(* Logix 5000 project; controller TFF vendor 1 type 14 code 107 rev 34.11; software revision 34.03; part 25 of 36 *)
(* tags used below, declared in another part *)
   Address : DINT;   // Temp Address
   Index : DINT;   // Index
   PCV101_PID_Settings : INT;
   sBar1 : STRING5;
   sBar2 : STRING5;
   sBar3 : STRING5;
   AnalogOutput : AnalogOutput[25];   // Analog Output Array
   Concentration : Concentration;
   ControlLoop_FeedBagLevel : ALIAS FOR ControlLoop[2];   // Feed Bag Level Control Loop
   ControlLoop_FeedPump : ALIAS FOR ControlLoop[1];   // Feed Pump Control Loop
   ControlLoop_PCV101 : ALIAS FOR ControlLoop[5];   // PCV101 Control Loop
   ControlLoop_PCV101_5ms : ALIAS FOR ControlLoop[6];   // PCV101 Control Loop
   ControlLoop_PCV101_CV : REAL;   // Control Value
   ControlLoop_PCV101_RAMP_OUT : REAL;   // Ramp Output
   DerivedData : DerivedData;   // Derived data (user input and calculated values)
   Diafiltration : Diafiltration;
   DigitalOutput : BOOL[256];   // Digital Output Array these bits are sent to output cards.
   DigitalPoint : DigitalPoint[150];   // Digital Point Array
   DP : ALIAS FOR AnalogPoint[40];   // Differential Pressure
   DPAlarm : ALIAS FOR AlarmAnalog[40];   // Differential Pressure Alarm
   Drive : Drive[11];   // Drives Array
   FI001 : ALIAS FOR AnalogPoint[42];   // Feed Flow
   FI001Alarm : ALIAS FOR AlarmAnalog[42];   // Feed Flow Alarm
   FI003 : ALIAS FOR AnalogPoint[17];
   FI101 : ALIAS FOR AnalogPoint[2];   // Filtrate Flow
   FI401 : ALIAS FOR AnalogPoint[43];   // Transfer Pump Flow
   FI401Alarm : ALIAS FOR AlarmAnalog[43];   // Transfer Pump Flow Alarm
   FlowPath : FlowPath[64];   // Flow Path Array
   FlowPathControl : FlowPathControl;   // Flow Path Control
   FQ_Conc : ALIAS FOR Totalizer[0];   // Concentration Totalizer
   FQ_Diaf : ALIAS FOR Totalizer[1];   // DiafiltrationTotalizer
   LI001 : ALIAS FOR AnalogPoint[44];   // Feed Bag Volume
   Membrane_Data : Membrane_Data;   // Membrane Data
   NWP : ALIAS FOR AnalogPoint[45];   // Normalized Water Permeability
   Options : Options;   // Options List
   PCV101_Control : PCV_Control;   // PCV101 Control UDT
   PERM : ALIAS FOR AnalogPoint[46];   // Membrane Permeability
   Phase : Phases[6];   // Phase Control Array
   Phase0 : ALIAS FOR Phase[0];   // Phase 0
   PhaseTotalizer : PhaseTotalizer[18];   // Phase Totalizers Array
   PI001 : ALIAS FOR AnalogPoint[5];   // Feed Pressure
   PI002 : ALIAS FOR AnalogPoint[6];   // Retentate Pressure
   PI101 : ALIAS FOR AnalogPoint[7];   // Filtrate Pressure
   PI401 : ALIAS FOR AnalogPoint[8];   // Transfer Pump Pressure
   PipeAnimation : PipeAnimation;   // HMI Pipe Animation Array
   SIC001 : ALIAS FOR Drive[1];   // Feed Pump
   SIC001DF : ALIAS FOR DigitalPoint[8];   // Feed Pump Defect
   SIC002 : ALIAS FOR Drive[2];   // Transfer Pump
   SIC002DF : ALIAS FOR DigitalPoint[9];   // Transfer Pump Defect
   SysControl : SysControl;   // General system status and command
   ThisSystem : SystemType;
   TI001 : ALIAS FOR AnalogPoint[13];   // Feed Bag Temperature
   TMP : ALIAS FOR AnalogPoint[41];   // Trans-membrane Pressure
   TMPAlarm : ALIAS FOR AlarmAnalog[41];   // Trans-membrane Pressure Alarm
   Totalizer : Totalizers[20];   // Totalizers Array
   XS011 : ALIAS FOR DigitalPoint[11];   // Pump P001 Type
   XS012 : ALIAS FOR DigitalPoint[12];   // Pump P002 Type
(* Process, continued *)

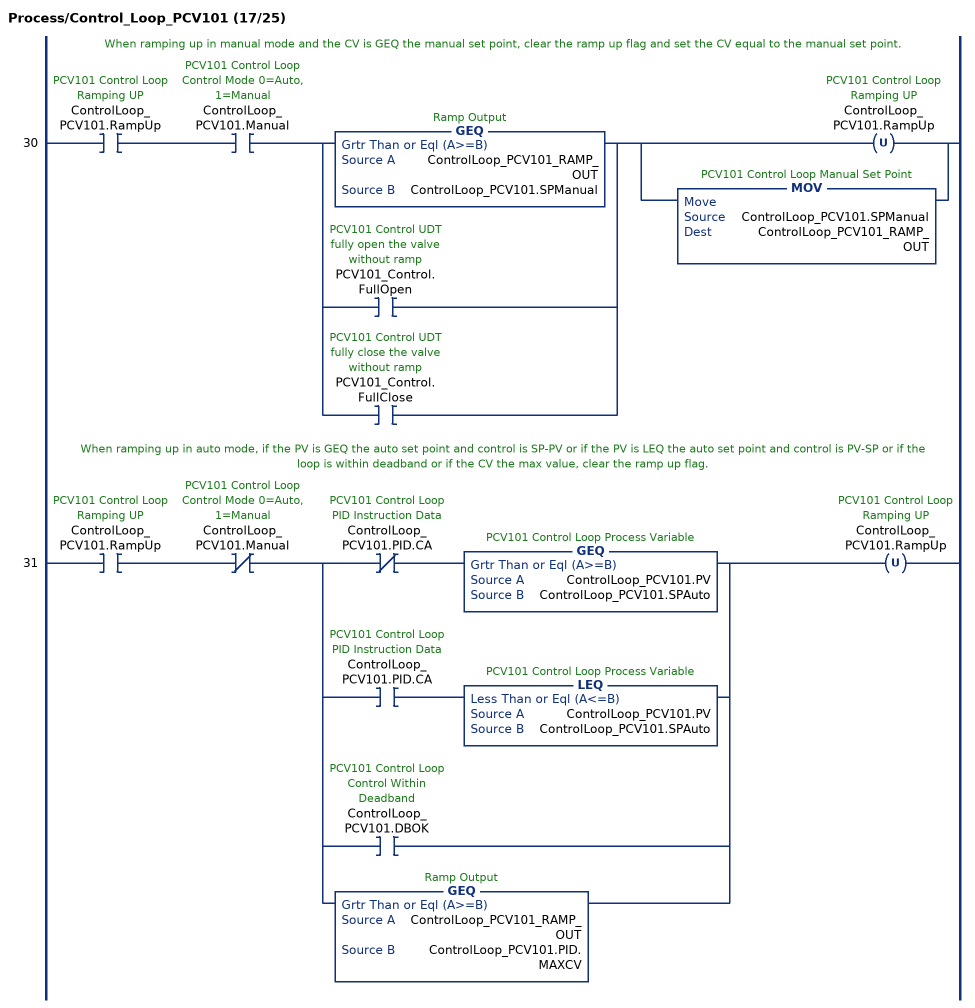
   [picture p237: Process/Control_Loop_PCV101 rungs 30-31]
   // When ramping up in manual mode and the CV is GEQ the manual set point, clear the ramp up flag and set the CV equal to the manual set point.
   30: XIC(ControlLoop_PCV101.RampUp)XIC(ControlLoop_PCV101.Manual)[GEQ(ControlLoop_PCV101_RAMP_OUT,ControlLoop_PCV101.SPManual) ,XIC(PCV101_Control.FullOpen) ,XIC(PCV101_Control.FullClose) ][OTU(ControlLoop_PCV101.RampUp) ,MOV(ControlLoop_PCV101.SPManual,ControlLoop_PCV101_RAMP_OUT) ];
   // When ramping up in auto mode, if the PV is GEQ the auto set point and control is SP-PV or if the PV is LEQ the auto set point and control is PV-SP or if the loop is within deadband or if the CV the max value, clear the ramp up flag.
   31: XIC(ControlLoop_PCV101.RampUp)XIO(ControlLoop_PCV101.Manual)[XIO(ControlLoop_PCV101.PID.CA) GEQ(ControlLoop_PCV101.PV,ControlLoop_PCV101.SPAuto) ,XIC(ControlLoop_PCV101.PID.CA) LEQ(ControlLoop_PCV101.PV,ControlLoop_PCV101.SPAuto) ,XIC(ControlLoop_PCV101.DBOK) ,GEQ(ControlLoop_PCV101_RAMP_OUT,ControlLoop_PCV101.PID.MAXCV) ]OTU(ControlLoop_PCV101.RampUp);
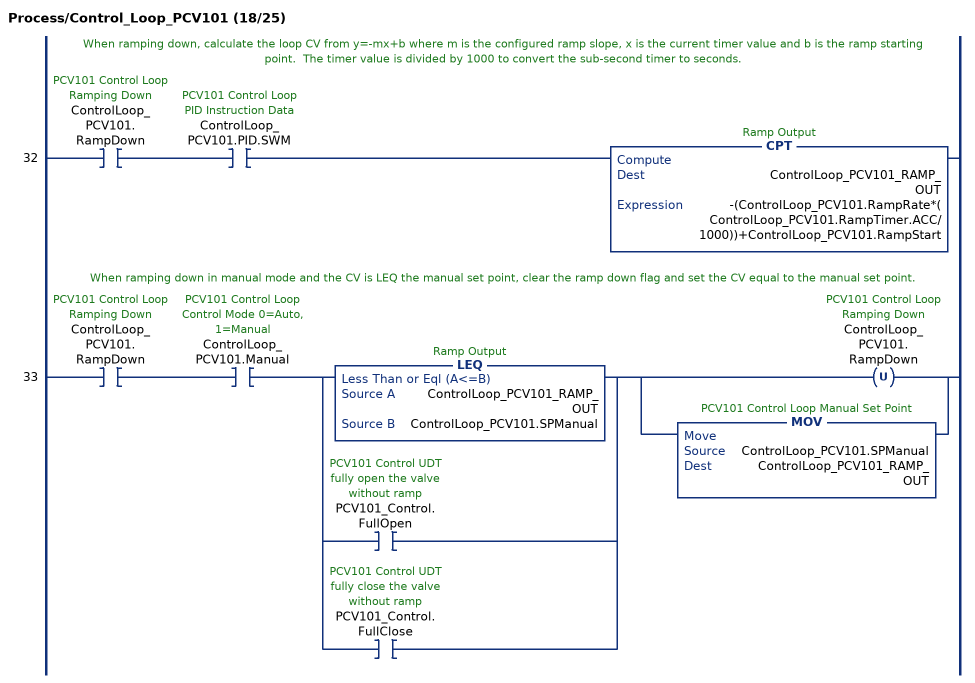
   // When ramping down, calculate the loop CV from y=-mx+b where m is the configured ramp slope, x is the current timer value and b is the ramp starting point.  The timer value is divided by 1000 to convert the sub-second timer to seconds.
   32: XIC(ControlLoop_PCV101.RampDown)XIC(ControlLoop_PCV101.PID.SWM)CPT(ControlLoop_PCV101_RAMP_OUT,-(ControlLoop_PCV101.RampRate*(ControlLoop_PCV101.RampTimer.ACC/1000))+ControlLoop_PCV101.RampStart);
   // When ramping down in manual mode and the CV is LEQ the manual set point, clear the ramp down flag and set the CV equal to the manual set point.
   33: XIC(ControlLoop_PCV101.RampDown)XIC(ControlLoop_PCV101.Manual)[LEQ(ControlLoop_PCV101_RAMP_OUT,ControlLoop_PCV101.SPManual) ,XIC(PCV101_Control.FullOpen) ,XIC(PCV101_Control.FullClose) ][OTU(ControlLoop_PCV101.RampDown) ,MOV(ControlLoop_PCV101.SPManual,ControlLoop_PCV101_RAMP_OUT) ];
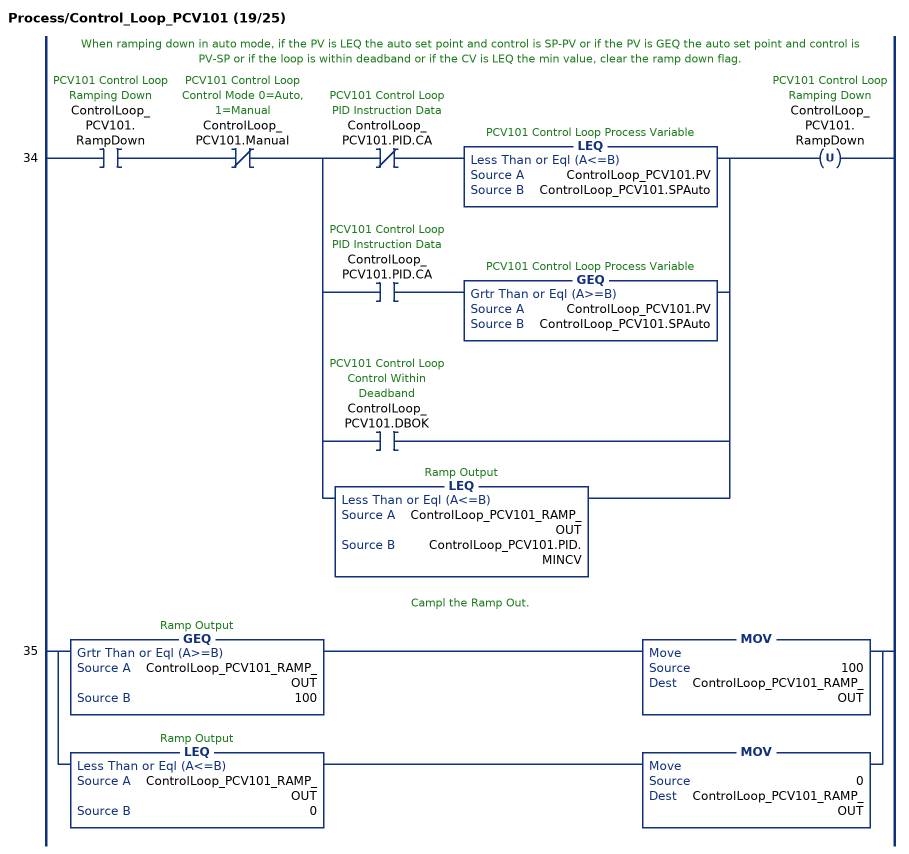
   // When ramping down in auto mode, if the PV is LEQ the auto set point and control is SP-PV or if the PV is GEQ the auto set point and control is PV-SP or if the loop is within deadband or if the CV is LEQ the min value, clear the ramp down flag.
   34: XIC(ControlLoop_PCV101.RampDown)XIO(ControlLoop_PCV101.Manual)[XIO(ControlLoop_PCV101.PID.CA) LEQ(ControlLoop_PCV101.PV,ControlLoop_PCV101.SPAuto) ,XIC(ControlLoop_PCV101.PID.CA) GEQ(ControlLoop_PCV101.PV,ControlLoop_PCV101.SPAuto) ,XIC(ControlLoop_PCV101.DBOK) ,LEQ(ControlLoop_PCV101_RAMP_OUT,ControlLoop_PCV101.PID.MINCV) ]OTU(ControlLoop_PCV101.RampDown);
   // Campl the Ramp Out.
   35: [GEQ(ControlLoop_PCV101_RAMP_OUT,100) MOV(100,ControlLoop_PCV101_RAMP_OUT) ,LEQ(ControlLoop_PCV101_RAMP_OUT,0) MOV(0,ControlLoop_PCV101_RAMP_OUT) ];
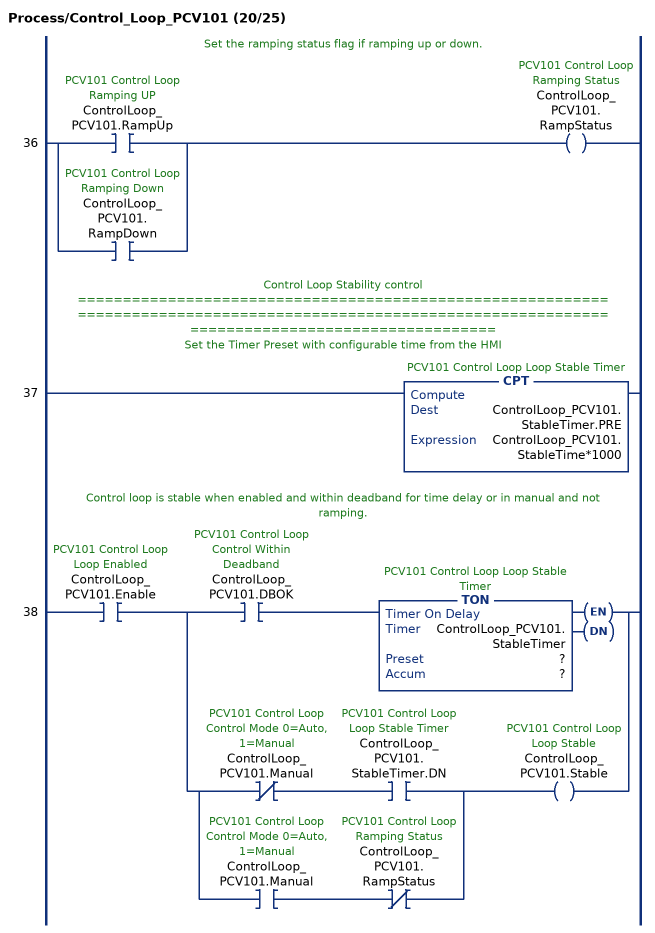
   // Set the ramping status flag if ramping up or down.
   36: [XIC(ControlLoop_PCV101.RampUp) ,XIC(ControlLoop_PCV101.RampDown) ]OTE(ControlLoop_PCV101.RampStatus);
   // Control Loop Stability control
   // ========================================================================================================================================================
   // Set the Timer Preset with configurable time from the HMI
   37: CPT(ControlLoop_PCV101.StableTimer.PRE,ControlLoop_PCV101.StableTime*1000);
   // Control loop is stable when enabled and within deadband for time delay or in manual and not ramping.
   38: XIC(ControlLoop_PCV101.Enable)[XIC(ControlLoop_PCV101.DBOK) TON(ControlLoop_PCV101.StableTimer,?,?) ,[XIO(ControlLoop_PCV101.Manual) XIC(ControlLoop_PCV101.StableTimer.DN) ,XIC(ControlLoop_PCV101.Manual) XIO(ControlLoop_PCV101.RampStatus) ] OTE(ControlLoop_PCV101.Stable) ];
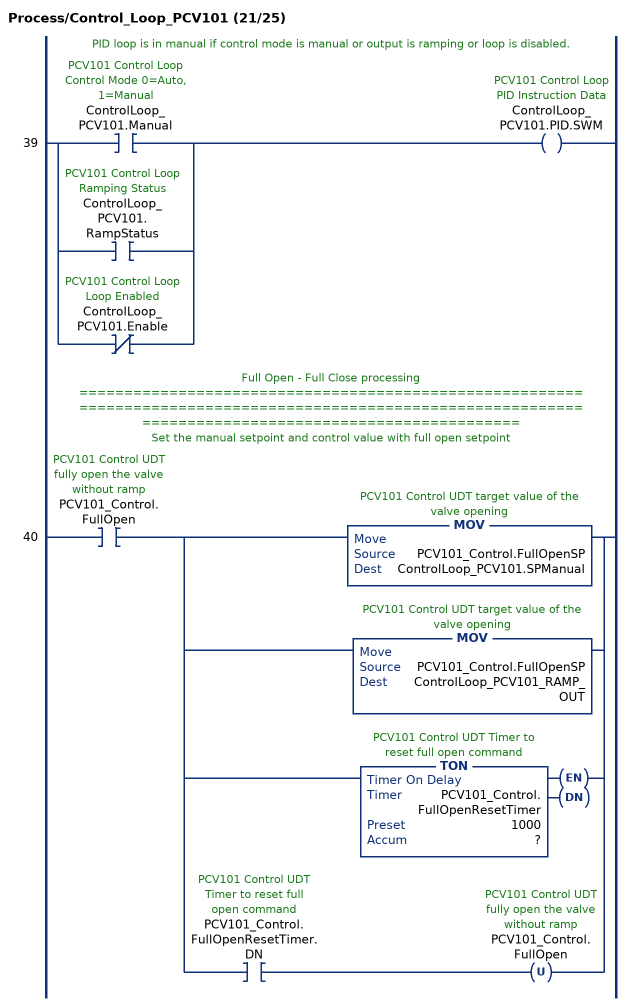
   // PID loop is in manual if control mode is manual or output is ramping or loop is disabled.
   39: [XIC(ControlLoop_PCV101.Manual) ,XIC(ControlLoop_PCV101.RampStatus) ,XIO(ControlLoop_PCV101.Enable) ]OTE(ControlLoop_PCV101.PID.SWM);
   // Full Open - Full Close processing
   // ==========================================================================================================================================================
   // Set the manual setpoint and control value with full open setpoint
   40: XIC(PCV101_Control.FullOpen)[MOV(PCV101_Control.FullOpenSP,ControlLoop_PCV101.SPManual) ,MOV(PCV101_Control.FullOpenSP,ControlLoop_PCV101_RAMP_OUT) ,TON(PCV101_Control.FullOpenResetTimer,?,?) ,XIC(PCV101_Control.FullOpenResetTimer.DN) OTU(PCV101_Control.FullOpen) ];
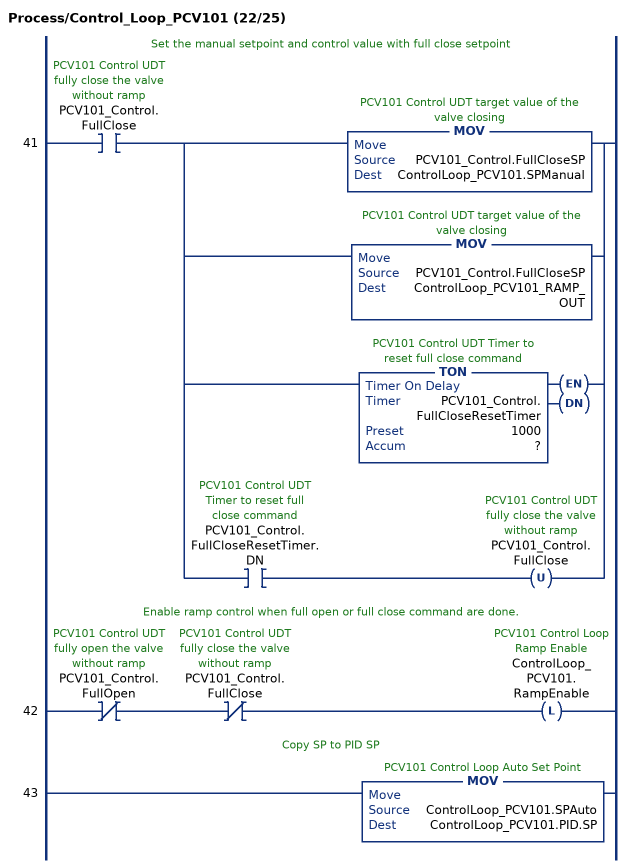
   // Set the manual setpoint and control value with full close setpoint
   41: XIC(PCV101_Control.FullClose)[MOV(PCV101_Control.FullCloseSP,ControlLoop_PCV101.SPManual) ,MOV(PCV101_Control.FullCloseSP,ControlLoop_PCV101_RAMP_OUT) ,TON(PCV101_Control.FullCloseResetTimer,?,?) ,XIC(PCV101_Control.FullCloseResetTimer.DN) OTU(PCV101_Control.FullClose) ];
   // Enable ramp control when full open or full close command are done.
   42: XIO(PCV101_Control.FullOpen)XIO(PCV101_Control.FullClose)OTL(ControlLoop_PCV101.RampEnable);
   // Copy SP to PID SP
   43: MOV(ControlLoop_PCV101.SPAuto,ControlLoop_PCV101.PID.SP);
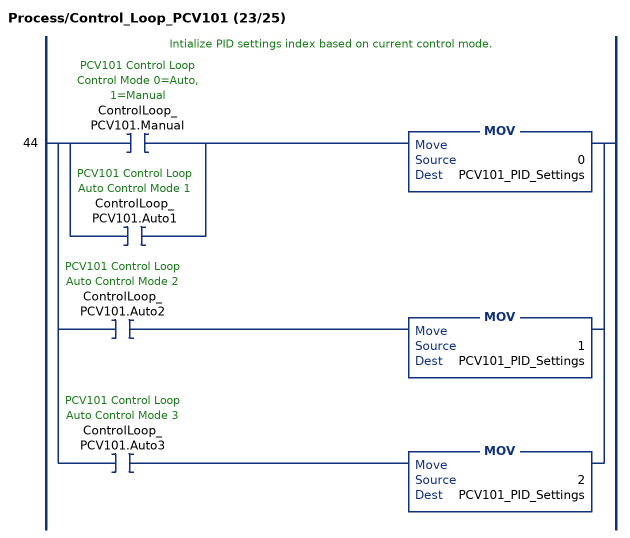
   // Intialize PID settings index based on current control mode.
   44: [[XIC(ControlLoop_PCV101.Manual) ,XIC(ControlLoop_PCV101.Auto1) ] MOV(0,PCV101_PID_Settings) ,XIC(ControlLoop_PCV101.Auto2) MOV(1,PCV101_PID_Settings) ,XIC(ControlLoop_PCV101.Auto3) MOV(2,PCV101_PID_Settings) ];
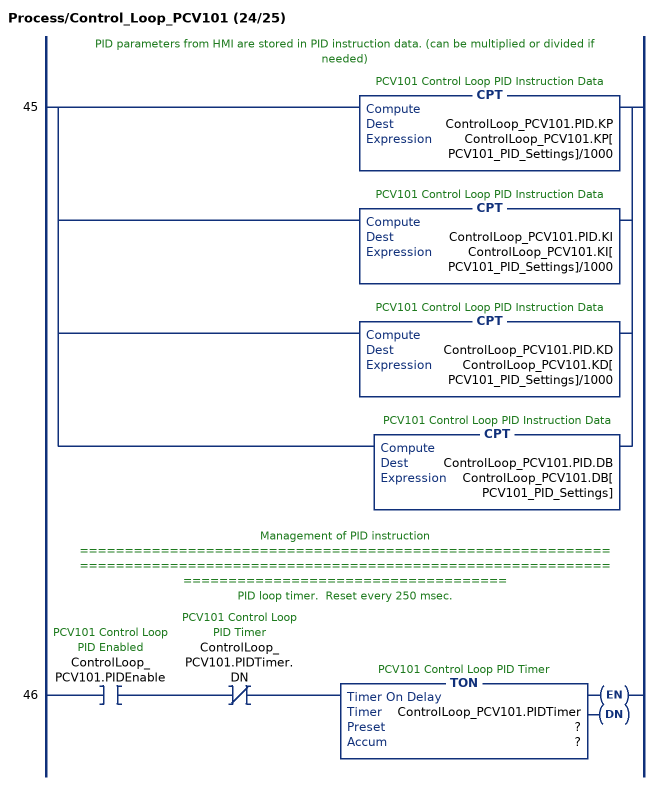
   // PID parameters from HMI are stored in PID instruction data. (can be multiplied or divided if needed)
   45: [CPT(ControlLoop_PCV101.PID.KP,ControlLoop_PCV101.KP[PCV101_PID_Settings]/1000) ,CPT(ControlLoop_PCV101.PID.KI,ControlLoop_PCV101.KI[PCV101_PID_Settings]/1000) ,CPT(ControlLoop_PCV101.PID.KD,ControlLoop_PCV101.KD[PCV101_PID_Settings]/1000) ,CPT(ControlLoop_PCV101.PID.DB,ControlLoop_PCV101.DB[PCV101_PID_Settings]) ];
   // Management of PID instruction
   // ==========================================================================================================================================================
   // PID loop timer.  Reset every 250 msec.
   46: XIC(ControlLoop_PCV101.PIDEnable)XIO(ControlLoop_PCV101.PIDTimer.DN)TON(ControlLoop_PCV101.PIDTimer,?,?);
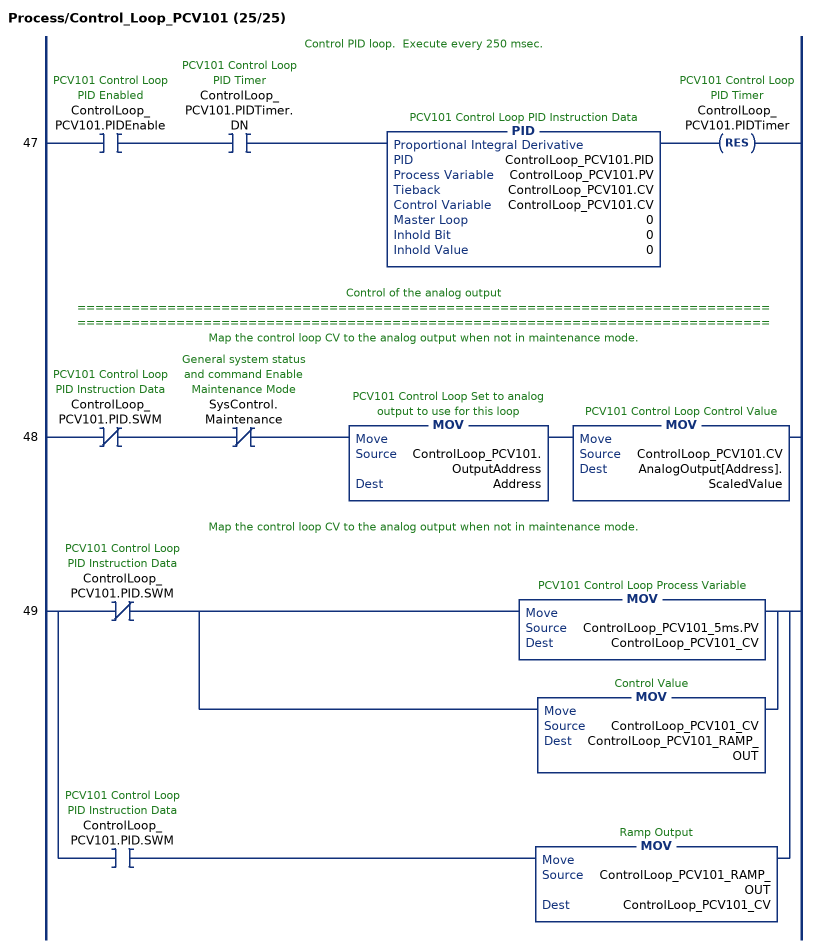
   // Control PID loop.  Execute every 250 msec.
   47: XIC(ControlLoop_PCV101.PIDEnable)XIC(ControlLoop_PCV101.PIDTimer.DN)PID(ControlLoop_PCV101.PID,ControlLoop_PCV101.PV,ControlLoop_PCV101.CV,ControlLoop_PCV101.CV,0,0,0)RES(ControlLoop_PCV101.PIDTimer);
   // Control of the analog output
   // ==========================================================================================================================================================
   // Map the control loop CV to the analog output when not in maintenance mode.
   48: XIO(ControlLoop_PCV101.PID.SWM)XIO(SysControl.Maintenance)MOV(ControlLoop_PCV101.OutputAddress,Address)MOV(ControlLoop_PCV101.CV,AnalogOutput[Address].ScaledValue);
   // Map the control loop CV to the analog output when not in maintenance mode.
   49: [XIO(ControlLoop_PCV101.PID.SWM) [MOV(ControlLoop_PCV101_5ms.PV,ControlLoop_PCV101_CV) ,MOV(ControlLoop_PCV101_CV,ControlLoop_PCV101_RAMP_OUT) ] ,XIC(ControlLoop_PCV101.PID.SWM) MOV(ControlLoop_PCV101_RAMP_OUT,ControlLoop_PCV101_CV) ];
END_ROUTINE

ROUTINE Derived_Data   (* structured text *)
// Derived Data Routine
   
   (* =======================================================================
   	Derived Data : calculations of derived data
   
   	List of treatments
   		- Derived Data Calculation
   
   -----------------------------------------------------------------------------------------------------------------------------------------------------
   	History
   		2019-AUG-13 - ACTEMIUM - B. Roch - Initial version for Candidate Release 3.00.00.00.a
   		2020-SEP-29 - Merck - Q. Spindler - Modifications for Candidate Release 3.00.00.01.a
   					- Add Retentate totalizers
   		2020-NOV-24 - Merck - Q. Spindler - Modifications for Candidate Release 3.00.00.01.b
   					- Change Retentate totalizers option
   =============================================================================================================================*)
   
   
   (* Derived Data Calculation
   =============================================================================================================================*)
   
   
   (* Compute pressure in PSI*)
   //Check Pressure at Feed Pump
   IF PI001.CurrentValue <= 0.00 Then
   	DerivedData.PI001_PSI := 0.00;
   ELSE
   //Check for bar vs. psig
   	IF PI001.EGU = sBar1 OR PI001.EGU = sBar2 OR PI001.EGU = sBar3 THEN
   		DerivedData.PI001_PSI := PI001.CurrentValue * 14.5;
   	ELSE;
   		DerivedData.PI001_PSI := PI001.CurrentValue;
   	END_IF;
   END_IF;
   //Check Pressure at Transfer Pump
   IF PI401.CurrentValue <= 0 Then
   	DerivedData.PI401_PSI:= 0.00;
   ELSE
   	//Check for bar vs. psig
   	IF PI401.EGU = sBar1 OR PI401.EGU = sBar2 OR PI401.EGU = sBar3 THEN
   		DerivedData.PI401_PSI := PI401.CurrentValue * 14.5;
   	ELSE;
   		DerivedData.PI401_PSI := PI401.CurrentValue;
   	END_IF;
   END_IF;
   
   
   (* Feed Flow Calculation*)
   IF Not SysControl.Simulate THEN
   	//If Pump is not running set flow to 0
   	IF NOT SIC001.RunStatus THEN;
   		FI001.CurrentValue := 0.0;
   	ELSE
   		IF ThisSystem.MoldType  = 124 THEN; // TF-3S system
   			IF Not FlowPathControl.FlushMode_Enabled THEN // NOT FLUSH MODE
   			FI001.CurrentValue := ((ControlLoop_FeedPump.CV - ((-0.00004*DerivedData.PI001_PSI*DerivedData.PI001_PSI*DerivedData.PI001_PSI) + (0.005*DerivedData.PI001_PSI*DerivedData.PI001_PSI) - (0.1725*DerivedData.PI001_PSI) + 0.2266)) / ((-0.00000002*DerivedData.PI001_PSI*DerivedData.PI001_PSI) + (0.000006*DerivedData.PI001_PSI) + 0.0012)) / 1000 ;
   			ELSE
   				IF DerivedData.PI001_PSI < 15 THEN FI001.CurrentValue := (0.00007*ControlLoop_FeedPump.CV*ControlLoop_FeedPump.CV*ControlLoop_FeedPump.CV) - (0.0125*ControlLoop_FeedPump.CV*ControlLoop_FeedPump.CV) + (0.8919*ControlLoop_FeedPump.CV+0.1849);
   				ELSE;
   					IF DerivedData.PI001_PSI < 25 THEN FI001.CurrentValue:=(-0.000009*ControlLoop_FeedPump.CV*ControlLoop_FeedPump.CV*ControlLoop_FeedPump.CV*ControlLoop_FeedPump.CV)+(0.0009*ControlLoop_FeedPump.CV*ControlLoop_FeedPump.CV*ControlLoop_FeedPump.CV)-(0.0349*ControlLoop_FeedPump.CV*ControlLoop_FeedPump.CV)+(1.0499*ControlLoop_FeedPump.CV);
   					ELSE;
   						IF DerivedData.PI001_PSI < 35 THEN FI001.CurrentValue:=(-0.0071*ControlLoop_FeedPump.CV*ControlLoop_FeedPump.CV)+(0.7692*ControlLoop_FeedPump.CV);
   						ELSE;
   							IF DerivedData.PI001_PSI < 50 THEN FI001.CurrentValue:=(0.0001*ControlLoop_FeedPump.CV*ControlLoop_FeedPump.CV*ControlLoop_FeedPump.CV)-(0.0135*ControlLoop_FeedPump.CV*ControlLoop_FeedPump.CV)+(0.8337*ControlLoop_FeedPump.CV);
   							ELSE FI001.CurrentValue:=(0.0001*ControlLoop_FeedPump.CV*ControlLoop_FeedPump.CV*ControlLoop_FeedPump.CV)-(0.0126*ControlLoop_FeedPump.CV*ControlLoop_FeedPump.CV)+(0.8045*ControlLoop_FeedPump.CV);
   							END_IF;
   						END_IF;
   					END_IF;
   				END_IF;
   			END_IF;
   		ELSE	// TF-2S system
   			// Check XS011 - Feed Pump type (0=1200S ; 1=150S)
   			IF Not(XS011.CurrentValue) THEN;
   				// 1200S :
   				FI001.CurrentValue := ControlLoop_FeedPump.CV / (4.3979 - (0.001788 * DerivedData.PI001_PSI) + (0.000495 * DerivedData.PI001_PSI * DerivedData.PI001_PSI) - (0.000005 * DerivedData.PI001_PSI * DerivedData.PI001_PSI * DerivedData.PI001_PSI)) ;
   			ELSE
   				// 150S :
   				FI001.CurrentValue := ControlLoop_FeedPump.CV / (4.3979 - (0.001788 * DerivedData.PI001_PSI) + (0.000495 * DerivedData.PI001_PSI * DerivedData.PI001_PSI) - (0.000005 * DerivedData.PI001_PSI * DerivedData.PI001_PSI * DerivedData.PI001_PSI)) ;
   			END_IF;
   		END_IF;
   	END_IF;
   END_IF;
   
   //Set flow to 0 if negative
   IF FI001.CurrentValue < 0 THEN FI001.CurrentValue := 0; END_IF;
   FI001Alarm.PV := FI001.CurrentValue;
   
   
   
   (* Transfer Flow Calculation*)
   IF Not SysControl.Simulate THEN
   	//If Pump is not running set flow to 0
   	IF NOT SIC002.RunStatus THEN;
   		FI401.CurrentValue := 0.0;
   	ELSE
   		IF ThisSystem.MoldType  = 124 THEN; // TF-3S system
   		FI401.CurrentValue := ControlLoop_FeedBagLevel.CV / (4.3979 - (0.001788 * DerivedData.PI401_PSI) + (0.000495 * DerivedData.PI401_PSI * DerivedData.PI401_PSI) - (0.000005 * DerivedData.PI401_PSI * DerivedData.PI401_PSI * DerivedData.PI401_PSI)) ;
   		ELSE	// TF-2S system
   			// Check XS012 - Transfer Pump type (0=1200S ; 1=150S)
   			IF Not(XS012.CurrentValue) THEN;
   				// 1200S :
   				FI401.CurrentValue := ControlLoop_FeedBagLevel.CV / (4.3979 - (0.001788 * DerivedData.PI401_PSI) + (0.000495 * DerivedData.PI401_PSI * DerivedData.PI401_PSI) - (0.000005 * DerivedData.PI401_PSI * DerivedData.PI401_PSI * DerivedData.PI401_PSI)) ;
   			ELSE
   				// 150S :
   				FI401.CurrentValue := ControlLoop_FeedBagLevel.CV / (4.3979 - (0.001788 * DerivedData.PI401_PSI) + (0.000495 * DerivedData.PI401_PSI * DerivedData.PI401_PSI) - (0.000005 * DerivedData.PI401_PSI * DerivedData.PI401_PSI * DerivedData.PI401_PSI)) ;
   			END_IF;
   		END_IF;
   	END_IF;
   END_IF;
   
   //Set flow to 0 if negative
   IF FI401.CurrentValue < 0 THEN FI401.CurrentValue := 0; END_IF;
   FI401Alarm.PV := FI401.CurrentValue;
   
   
   
   (*Differential Pressure*)
   DP.CurrentValue := PI001.CurrentValue - PI002.CurrentValue;
   DPAlarm.PV := DP.CurrentValue;
   
   
   (*Trans-Membrane Pressure*)
   TMP.CurrentValue := ((PI001.CurrentValue + PI002.CurrentValue) / 2) - PI101.CurrentValue;
   TMPAlarm.PV := TMP.CurrentValue;
   
   
   (*Flux : Membrane Flux*)
   Membrane_Data.Flux := FI101.CurrentValue / Membrane_Data.Area * 60;
   
   (*Diafiltration Volumes*)
   Diafiltration.Diaf_Volume := FQ_Diaf.Total / (Diafiltration.Diaf_Init + DerivedData.HOLDUP);
   
   (*VCF : Volume Concentration Factor*)
   Concentration.VCF := (LI001.CurrentValue + FQ_Conc.Total) / (LI001.CurrentValue + DerivedData.HOLDUP);
   
   (*Clamp VCF Value if less than 1*)
   IF Concentration.VCF < 1 THEN Concentration.VCF := 1; END_IF;
   
   (*CB : Protein Concentration*)
   Concentration.CB := Concentration.Conc_Init * Concentration.VCF;
   
   
   (*NWP TCF*)
   
   (*Fill Lookup Table for TCF 25 DegC*)
   Membrane_Data.NWP_TCF_Lookup_25[0] := 2.011;
   Membrane_Data.NWP_TCF_Lookup_25[1] := 1.943;
   Membrane_Data.NWP_TCF_Lookup_25[2] := 1.879;
   Membrane_Data.NWP_TCF_Lookup_25[3] := 1.818;
   Membrane_Data.NWP_TCF_Lookup_25[4] := 1.761;
   Membrane_Data.NWP_TCF_Lookup_25[5] := 1.706;
   Membrane_Data.NWP_TCF_Lookup_25[6] := 1.653;
   Membrane_Data.NWP_TCF_Lookup_25[7] := 1.604;
   Membrane_Data.NWP_TCF_Lookup_25[8] := 1.556;
   Membrane_Data.NWP_TCF_Lookup_25[9] := 1.511;
   Membrane_Data.NWP_TCF_Lookup_25[10] := 1.468;
   Membrane_Data.NWP_TCF_Lookup_25[11] := 1.426;
   Membrane_Data.NWP_TCF_Lookup_25[12] := 1.387;
   Membrane_Data.NWP_TCF_Lookup_25[13] := 1.349;
   Membrane_Data.NWP_TCF_Lookup_25[14] := 1.313;
   Membrane_Data.NWP_TCF_Lookup_25[15] := 1.278;
   Membrane_Data.NWP_TCF_Lookup_25[16] := 1.245;
   Membrane_Data.NWP_TCF_Lookup_25[17] := 1.213;
   Membrane_Data.NWP_TCF_Lookup_25[18] := 1.183;
   Membrane_Data.NWP_TCF_Lookup_25[19] := 1.154;
   Membrane_Data.NWP_TCF_Lookup_25[20] := 1.126;
   Membrane_Data.NWP_TCF_Lookup_25[21] := 1.099;
   Membrane_Data.NWP_TCF_Lookup_25[22] := 1.072;
   Membrane_Data.NWP_TCF_Lookup_25[23] := 1.047;
   Membrane_Data.NWP_TCF_Lookup_25[24] := 1.022;
   Membrane_Data.NWP_TCF_Lookup_25[25] := 1.0;
   Membrane_Data.NWP_TCF_Lookup_25[26] := 0.978;
   Membrane_Data.NWP_TCF_Lookup_25[27] := 0.956;
   Membrane_Data.NWP_TCF_Lookup_25[28] := 0.935;
   Membrane_Data.NWP_TCF_Lookup_25[29] := 0.915;
   Membrane_Data.NWP_TCF_Lookup_25[30] := 0.896;
   Membrane_Data.NWP_TCF_Lookup_25[31] := 0.877;
   Membrane_Data.NWP_TCF_Lookup_25[32] := 0.859;
   Membrane_Data.NWP_TCF_Lookup_25[33] := 0.841;
   Membrane_Data.NWP_TCF_Lookup_25[34] := 0.824;
   Membrane_Data.NWP_TCF_Lookup_25[35] := 0.808;
   Membrane_Data.NWP_TCF_Lookup_25[36] := 0.791;
   Membrane_Data.NWP_TCF_Lookup_25[37] := 0.777;
   Membrane_Data.NWP_TCF_Lookup_25[38] := 0.761;
   Membrane_Data.NWP_TCF_Lookup_25[39] := 0.747;
   Membrane_Data.NWP_TCF_Lookup_25[40] := 0.733;
   Membrane_Data.NWP_TCF_Lookup_25[41] := 0.719;
   Membrane_Data.NWP_TCF_Lookup_25[42] := 0.706;
   Membrane_Data.NWP_TCF_Lookup_25[43] := 0.694;
   Membrane_Data.NWP_TCF_Lookup_25[44] := 0.681;
   Membrane_Data.NWP_TCF_Lookup_25[45] := 0.669;
   Membrane_Data.NWP_TCF_Lookup_25[46] := 0.658;
   Membrane_Data.NWP_TCF_Lookup_25[47] := 0.646;
   Membrane_Data.NWP_TCF_Lookup_25[48] := 0.635;
   Membrane_Data.NWP_TCF_Lookup_25[49] := 0.624;
   Membrane_Data.NWP_TCF_Lookup_25[50] := 0.614;
   Membrane_Data.NWP_TCF_Lookup_25[51] := 0.604;
   Membrane_Data.NWP_TCF_Lookup_25[52] := 0.594;
   
   (*Compute NWP_TCF based on Lookup Table for TCF 25 DegC*)
   IF TI001.CurrentValue < 0 THEN;
   	(*Temperature below lookup table values*)
   	Membrane_Data.NWP_TCF:= Membrane_Data.NWP_TCF_Lookup_25[0];
   ELSIF TI001.CurrentValue> 51 THEN;
   	(*Temperature above lookup table values*)
   	Membrane_Data.NWP_TCF:= Membrane_Data.NWP_TCF_Lookup_25[52];
   ELSE
   	(*Temperature within lookup table values*)
   	Membrane_Data.NWP_TCF_Temp:= TRUNC(TI001.CurrentValue);
   	Membrane_Data.NWP_TCF:= (TI001.CurrentValue-Membrane_Data.NWP_TCF_Temp) * ( Membrane_Data.NWP_TCF_Lookup_25[Membrane_Data.NWP_TCF_Temp+1] - Membrane_Data.NWP_TCF_Lookup_25[Membrane_Data.NWP_TCF_Temp] ) + Membrane_Data.NWP_TCF_Lookup_25[Membrane_Data.NWP_TCF_Temp];
   END_IF;
   
   
   (*NWP : Normalized Water Permeability*)
   IF TMP.CurrentValue <> 0 THEN NWP.CurrentValue := Membrane_Data.Flux * Membrane_Data.NWP_TCF / TMP.CurrentValue; ELSE NWP.CurrentValue := 0; END_IF;
   
   
   
   (*PERM : Membrane Permeability*)
   IF TMP.CurrentValue <> 0 THEN PERM.CurrentValue := Membrane_Data.Flux / TMP.CurrentValue; ELSE PERM.CurrentValue := 0; END_IF;
   
   
   (*Reset Filtrate totalizer if option is disabled*)
   IF Options.No_Filtrate_Measurement THEN
   	FOR Index := 6 TO 11 DO;
   		PhaseTotalizer[Index].Phase := 0;
   		PhaseTotalizer[Index].Step := 0;
   		PhaseTotalizer[Index].Pause := 0;
   		PhaseTotalizer[Index].User := 0;
   		PhaseTotalizer[Index].Procedure := 0;
   	END_FOR;
   END_IF;
   
   
   (*Reset Retentate totalizer if option is disabled*)
   IF not Options.FI003 THEN
   	FOR Index := 12 TO 17 DO;
   		PhaseTotalizer[Index].Phase := 0;
   		PhaseTotalizer[Index].Step := 0;
   		PhaseTotalizer[Index].Pause := 0;
   		PhaseTotalizer[Index].User := 0;
   		PhaseTotalizer[Index].Procedure := 0;
   	END_FOR;
   END_IF;
END_ROUTINE

ROUTINE Drive_SIC001_Feed   (* ladder *)
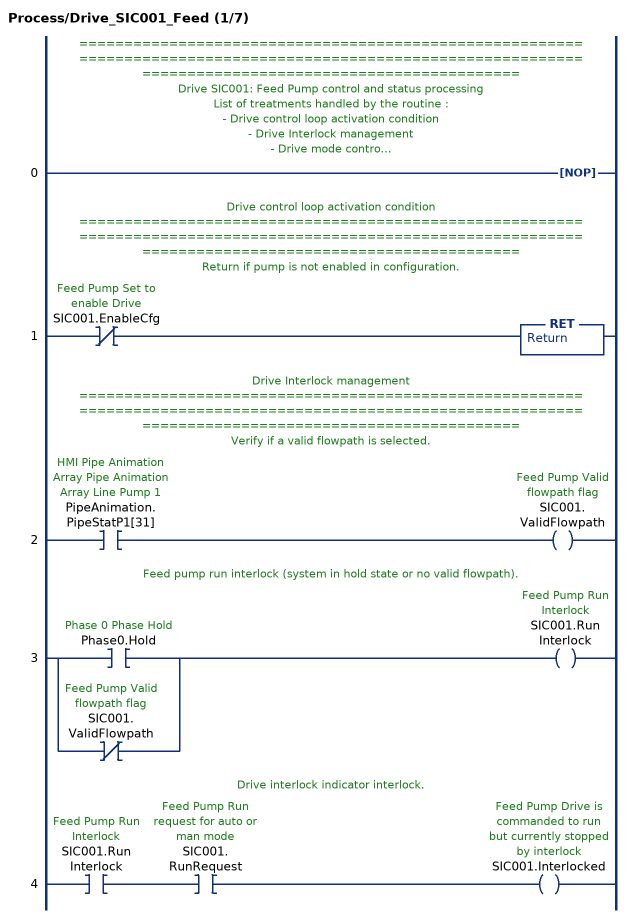
   // ==========================================================================================================================================================
   //                                                    Drive SIC001: Feed Pump control and status processing
   //                                                     List of treatments handled by the routine :
   //                                                          - Drive control loop activation condition
   //                                                          - Drive Interlock management
   //                                                          - Drive mode control
   //                                                          - Drive run command control
   //                                                          - Drive status management
   //                                                          - Drive status for HMI
   //                                                          - Drive DigitalOutput control
   //                                                     -----------------------------------------------------------------------------------------------------------------------------------------------------
   //                                                     History
   //                                                          2019-AUG-13 - Actemium - B. Roch - Initial version for Candidate Release 3.00.00.00.a
   // ==========================================================================================================================================================
   0: NOP();
   // Drive control loop activation condition
   // ==========================================================================================================================================================
   // Return if pump is not enabled in configuration.
   1: XIO(SIC001.EnableCfg)RET();
   // Drive Interlock management
   // ==========================================================================================================================================================
   // Verify if a valid flowpath is selected.
   2: XIC(PipeAnimation.PipeStatP1[31])OTE(SIC001.ValidFlowpath);
   // Feed pump run interlock (system in hold state or no valid flowpath).
   3: [XIC(Phase0.Hold) ,XIO(SIC001.ValidFlowpath) ]OTE(SIC001.RunInterlock);
   // Drive interlock indicator interlock.
   4: XIC(SIC001.RunInterlock)XIC(SIC001.RunRequest)OTE(SIC001.Interlocked);
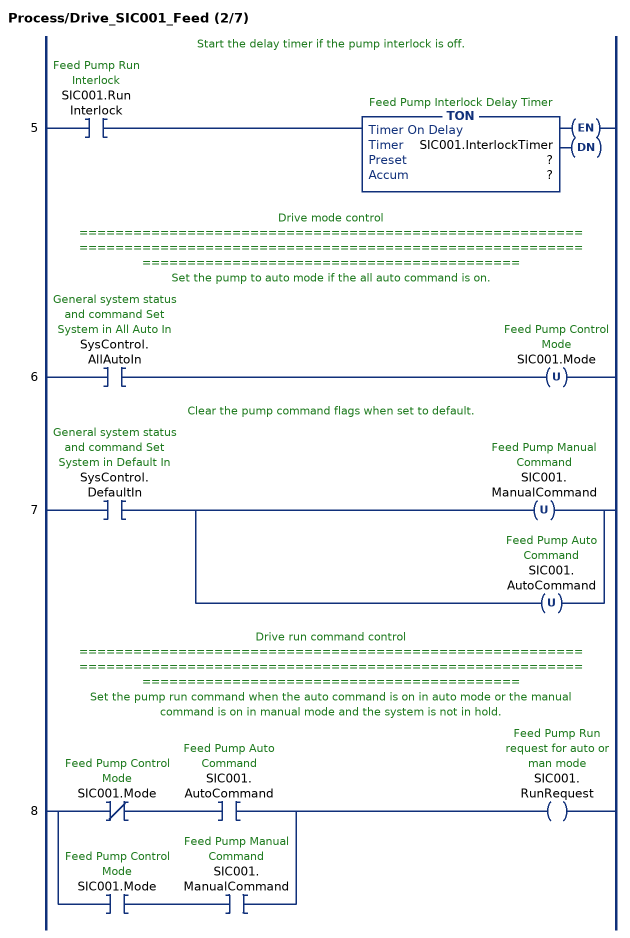
   // Start the delay timer if the pump interlock is off.
   5: XIC(SIC001.RunInterlock)TON(SIC001.InterlockTimer,?,?);
   // Drive mode control
   // ==========================================================================================================================================================
   // Set the pump to auto mode if the all auto command is on.
   6: XIC(SysControl.AllAutoIn)OTU(SIC001.Mode);
   // Clear the pump command flags when set to default.
   7: XIC(SysControl.DefaultIn)[OTU(SIC001.ManualCommand) ,OTU(SIC001.AutoCommand) ];
   // Drive run command control
   // ==========================================================================================================================================================
   // Set the pump run command when the auto command is on in auto mode or the manual command is on in manual mode and the system is not in hold.
   8: [XIO(SIC001.Mode) XIC(SIC001.AutoCommand) ,XIC(SIC001.Mode) XIC(SIC001.ManualCommand) ]OTE(SIC001.RunRequest);
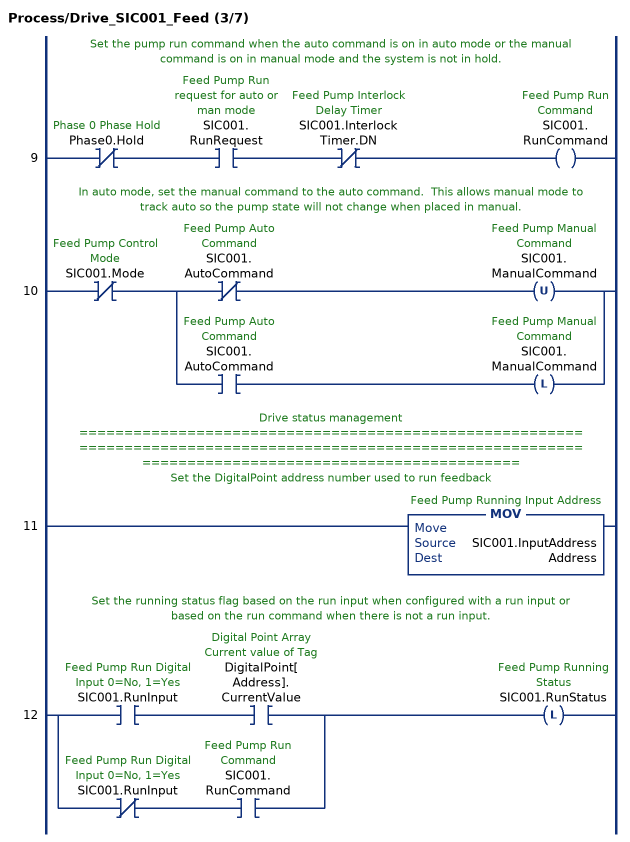
   // Set the pump run command when the auto command is on in auto mode or the manual command is on in manual mode and the system is not in hold.
   9: XIO(Phase0.Hold)XIC(SIC001.RunRequest)XIO(SIC001.InterlockTimer.DN)OTE(SIC001.RunCommand);
   // In auto mode, set the manual command to the auto command.  This allows manual mode to track auto so the pump state will not change when placed in manual.
   10: XIO(SIC001.Mode)[XIO(SIC001.AutoCommand) OTU(SIC001.ManualCommand) ,XIC(SIC001.AutoCommand) OTL(SIC001.ManualCommand) ];
   // Drive status management
   // ==========================================================================================================================================================
   // Set the DigitalPoint address number used to run feedback
   11: MOV(SIC001.InputAddress,Address);
   // Set the running status flag based on the run input when configured with a run input or based on the run command when there is not a run input.
   12: [XIC(SIC001.RunInput) XIC(DigitalPoint[Address].CurrentValue) ,XIO(SIC001.RunInput) XIC(SIC001.RunCommand) ]OTL(SIC001.RunStatus);
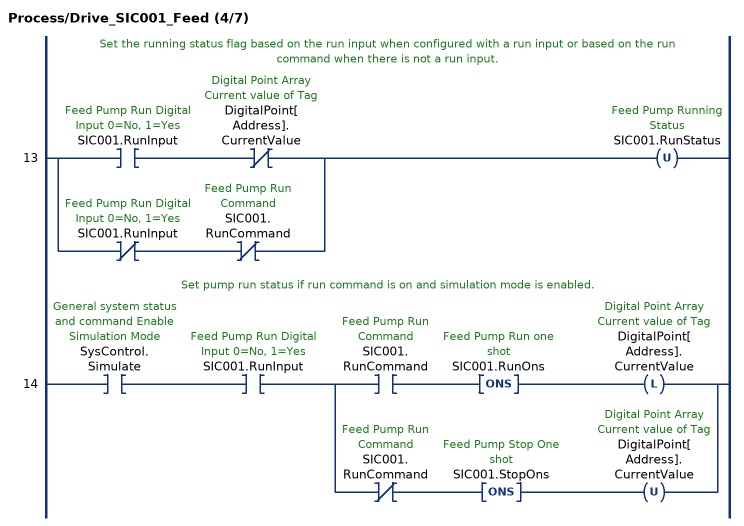
   // Set the running status flag based on the run input when configured with a run input or based on the run command when there is not a run input.
   13: [XIC(SIC001.RunInput) XIO(DigitalPoint[Address].CurrentValue) ,XIO(SIC001.RunInput) XIO(SIC001.RunCommand) ]OTU(SIC001.RunStatus);
   // Set pump run status if run command is on and simulation mode is enabled.
   14: XIC(SysControl.Simulate)XIC(SIC001.RunInput)[XIC(SIC001.RunCommand) ONS(SIC001.RunOns) OTL(DigitalPoint[Address].CurrentValue) ,XIO(SIC001.RunCommand) ONS(SIC001.StopOns) OTU(DigitalPoint[Address].CurrentValue) ];
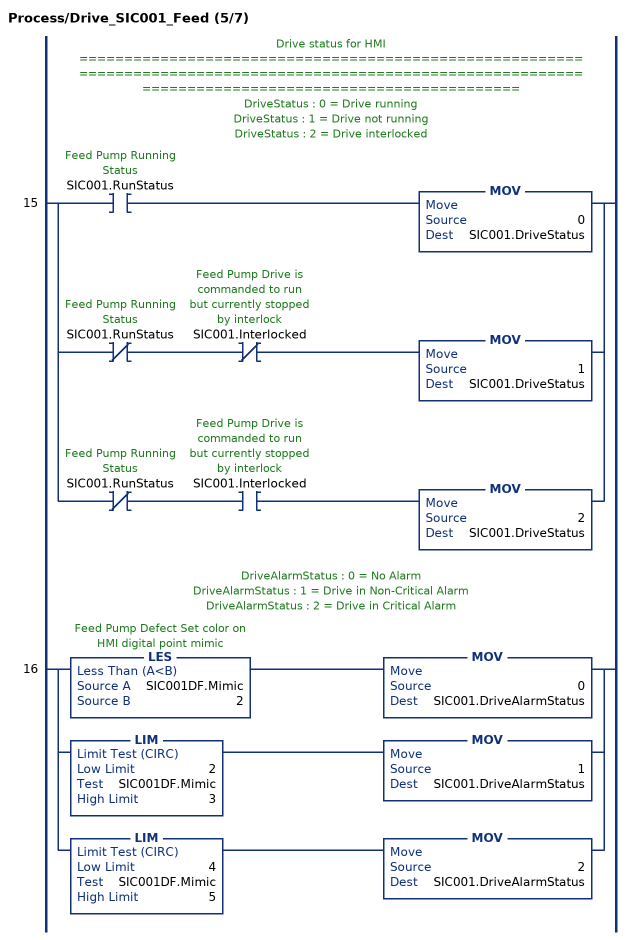
   // Drive status for HMI
   // ==========================================================================================================================================================
   //  DriveStatus : 0 = Drive running
   //  DriveStatus : 1 = Drive not running
   //  DriveStatus : 2 = Drive interlocked
   15: [XIC(SIC001.RunStatus) MOV(0,SIC001.DriveStatus) ,XIO(SIC001.RunStatus) XIO(SIC001.Interlocked) MOV(1,SIC001.DriveStatus) ,XIO(SIC001.RunStatus) XIC(SIC001.Interlocked) MOV(2,SIC001.DriveStatus) ];
   // DriveAlarmStatus : 0 = No Alarm
   //  DriveAlarmStatus : 1 = Drive in Non-Critical Alarm
   //  DriveAlarmStatus : 2 = Drive in Critical Alarm
   16: [LES(SIC001DF.Mimic,2) MOV(0,SIC001.DriveAlarmStatus) ,LIM(2,SIC001DF.Mimic,3) MOV(1,SIC001.DriveAlarmStatus) ,LIM(4,SIC001DF.Mimic,5) MOV(2,SIC001.DriveAlarmStatus) ];
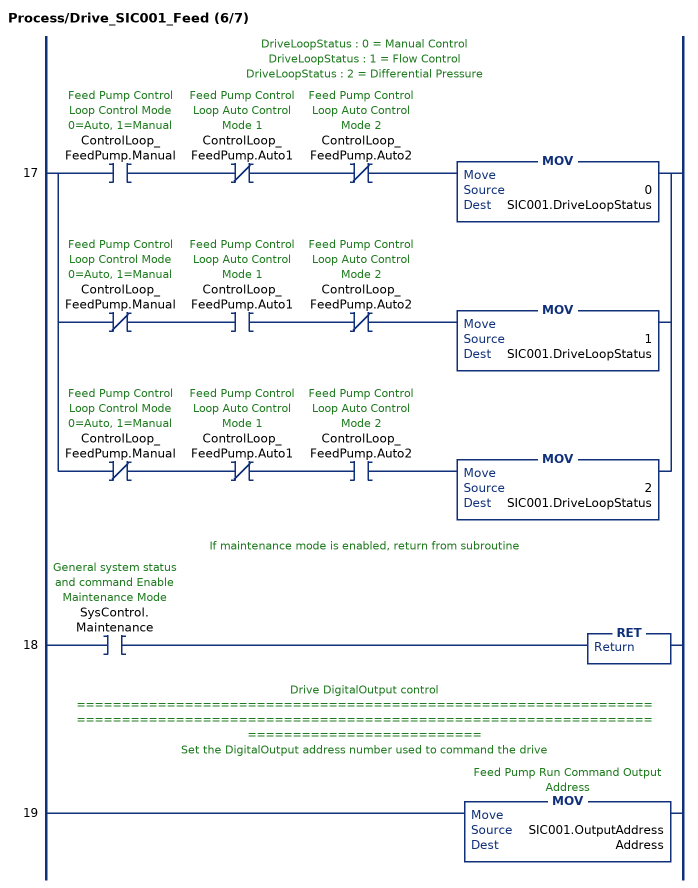
   // DriveLoopStatus : 0 = Manual Control
   //  DriveLoopStatus : 1 = Flow Control
   //  DriveLoopStatus : 2 = Differential Pressure
   17: [XIC(ControlLoop_FeedPump.Manual) XIO(ControlLoop_FeedPump.Auto1) XIO(ControlLoop_FeedPump.Auto2) MOV(0,SIC001.DriveLoopStatus) ,XIO(ControlLoop_FeedPump.Manual) XIC(ControlLoop_FeedPump.Auto1) XIO(ControlLoop_FeedPump.Auto2) MOV(1,SIC001.DriveLoopStatus) ,XIO(ControlLoop_FeedPump.Manual) XIO(ControlLoop_FeedPump.Auto1) XIC(ControlLoop_FeedPump.Auto2) MOV(2,SIC001.DriveLoopStatus) ];
   // If maintenance mode is enabled, return from subroutine
   18: XIC(SysControl.Maintenance)RET();
   // Drive DigitalOutput control
   // ==========================================================================================================================================================
   // Set the DigitalOutput address number used to command the drive
   19: MOV(SIC001.OutputAddress,Address);
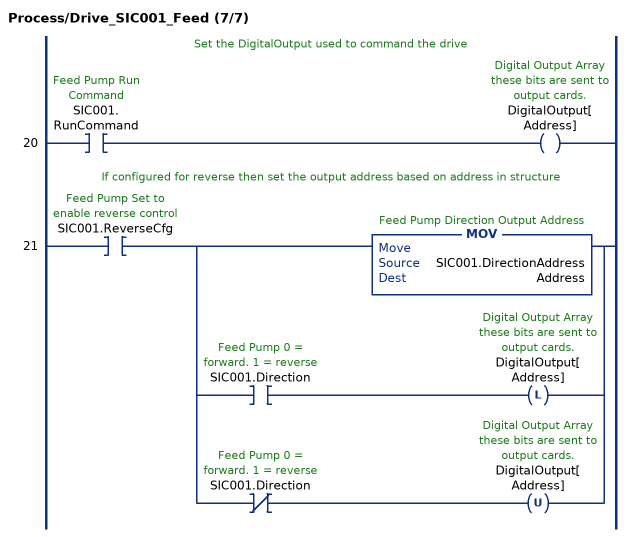
   // Set the DigitalOutput used to command the drive
   20: XIC(SIC001.RunCommand)OTE(DigitalOutput[Address]);
   // If configured for reverse then set the output address based on address in structure
   21: XIC(SIC001.ReverseCfg)[MOV(SIC001.DirectionAddress,Address) ,XIC(SIC001.Direction) OTL(DigitalOutput[Address]) ,XIO(SIC001.Direction) OTU(DigitalOutput[Address]) ];
END_ROUTINE

ROUTINE Drive_SIC002_Transfer   (* ladder *)
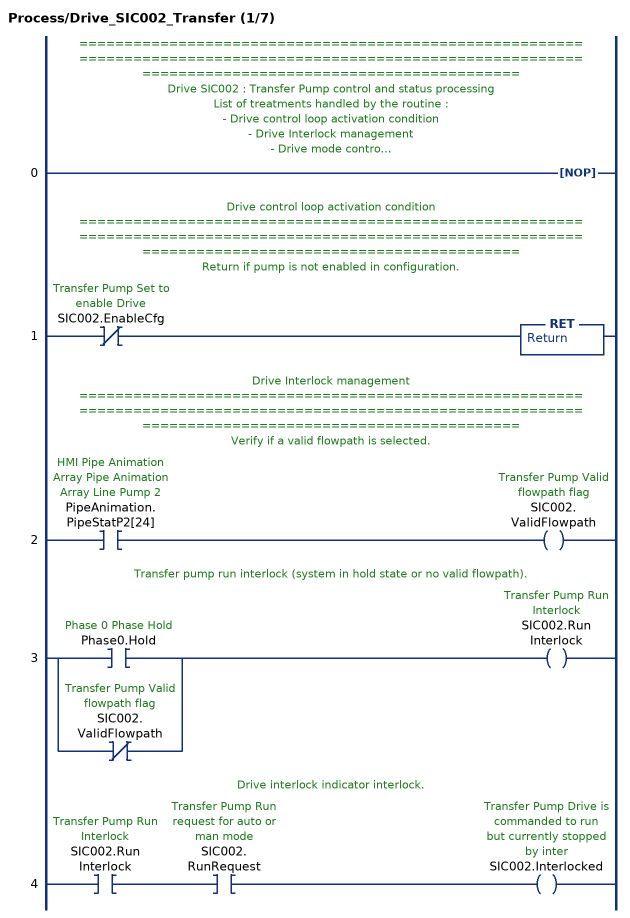
   // ==========================================================================================================================================================
   //                                                              Drive SIC002 : Transfer Pump control and status processing
   //                                                     List of treatments handled by the routine :
   //                                                          - Drive control loop activation condition
   //                                                          - Drive Interlock management
   //                                                          - Drive mode control
   //                                                          - Drive run command control
   //                                                          - Drive status management
   //                                                          - Drive status for HMI
   //                                                          - Drive DigitalOutput control
   //                                                     -----------------------------------------------------------------------------------------------------------------------------------------------------
   //                                                     History
   //                                                          2019-AUG-13 - Actemium - B. Roch - Initial version for Candidate Release 3.00.00.00.a
   // ==========================================================================================================================================================
   0: NOP();
   // Drive control loop activation condition
   // ==========================================================================================================================================================
   // Return if pump is not enabled in configuration.
   1: XIO(SIC002.EnableCfg)RET();
   // Drive Interlock management
   // ==========================================================================================================================================================
   // Verify if a valid flowpath is selected.
   2: XIC(PipeAnimation.PipeStatP2[24])OTE(SIC002.ValidFlowpath);
   // Transfer pump run interlock (system in hold state or no valid flowpath).
   3: [XIC(Phase0.Hold) ,XIO(SIC002.ValidFlowpath) ]OTE(SIC002.RunInterlock);
   // Drive interlock indicator interlock.
   4: XIC(SIC002.RunInterlock)XIC(SIC002.RunRequest)OTE(SIC002.Interlocked);
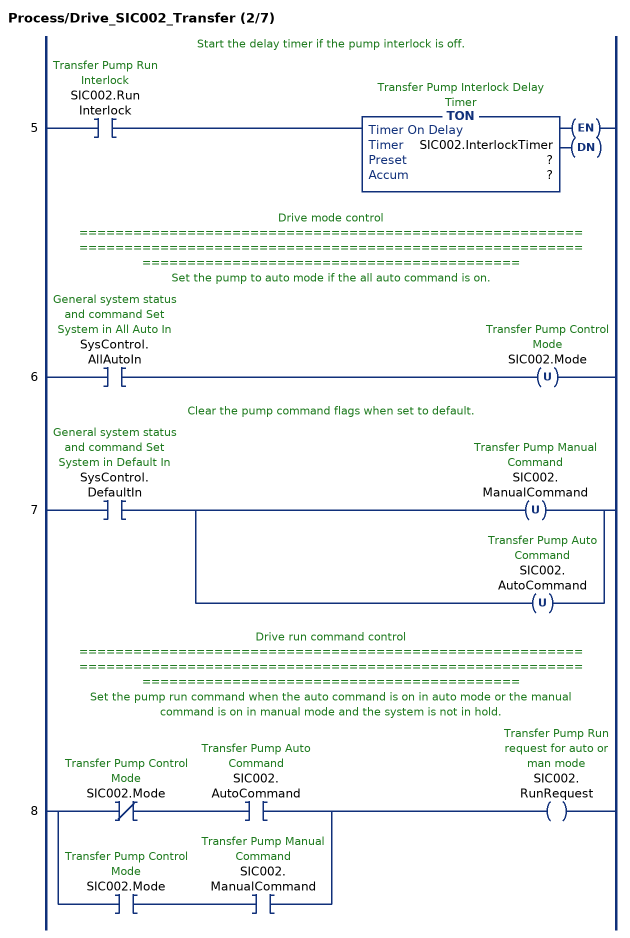
   // Start the delay timer if the pump interlock is off.
   5: XIC(SIC002.RunInterlock)TON(SIC002.InterlockTimer,?,?);
   // Drive mode control
   // ==========================================================================================================================================================
   // Set the pump to auto mode if the all auto command is on.
   6: XIC(SysControl.AllAutoIn)OTU(SIC002.Mode);
   // Clear the pump command flags when set to default.
   7: XIC(SysControl.DefaultIn)[OTU(SIC002.ManualCommand) ,OTU(SIC002.AutoCommand) ];
   // Drive run command control
   // ==========================================================================================================================================================
   // Set the pump run command when the auto command is on in auto mode or the manual command is on in manual mode and the system is not in hold.
   8: [XIO(SIC002.Mode) XIC(SIC002.AutoCommand) ,XIC(SIC002.Mode) XIC(SIC002.ManualCommand) ]OTE(SIC002.RunRequest);
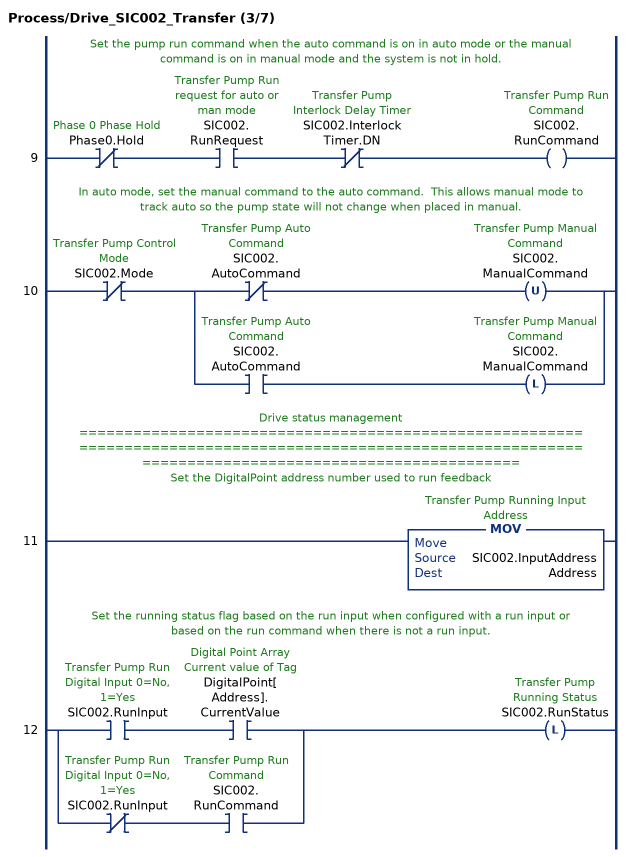
   // Set the pump run command when the auto command is on in auto mode or the manual command is on in manual mode and the system is not in hold.
   9: XIO(Phase0.Hold)XIC(SIC002.RunRequest)XIO(SIC002.InterlockTimer.DN)OTE(SIC002.RunCommand);
   // In auto mode, set the manual command to the auto command.  This allows manual mode to track auto so the pump state will not change when placed in manual.
   10: XIO(SIC002.Mode)[XIO(SIC002.AutoCommand) OTU(SIC002.ManualCommand) ,XIC(SIC002.AutoCommand) OTL(SIC002.ManualCommand) ];
   // Drive status management
   // ==========================================================================================================================================================
   // Set the DigitalPoint address number used to run feedback
   11: MOV(SIC002.InputAddress,Address);
   // Set the running status flag based on the run input when configured with a run input or based on the run command when there is not a run input.
   12: [XIC(SIC002.RunInput) XIC(DigitalPoint[Address].CurrentValue) ,XIO(SIC002.RunInput) XIC(SIC002.RunCommand) ]OTL(SIC002.RunStatus);
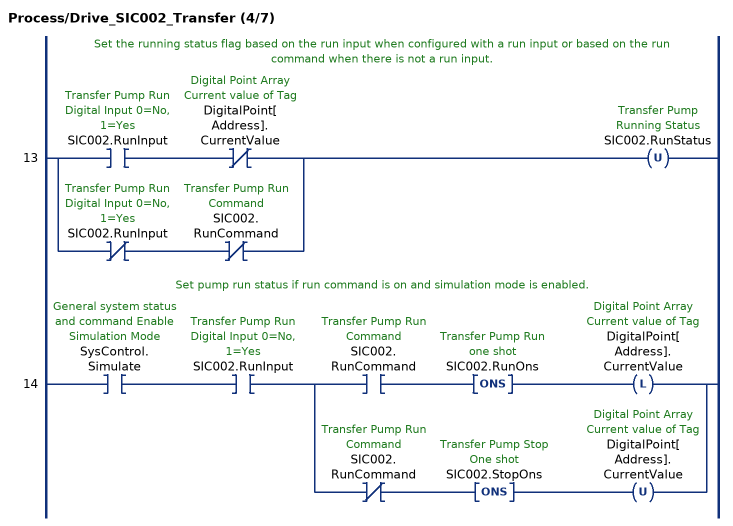
   // Set the running status flag based on the run input when configured with a run input or based on the run command when there is not a run input.
   13: [XIC(SIC002.RunInput) XIO(DigitalPoint[Address].CurrentValue) ,XIO(SIC002.RunInput) XIO(SIC002.RunCommand) ]OTU(SIC002.RunStatus);
   // Set pump run status if run command is on and simulation mode is enabled.
   14: XIC(SysControl.Simulate)XIC(SIC002.RunInput)[XIC(SIC002.RunCommand) ONS(SIC002.RunOns) OTL(DigitalPoint[Address].CurrentValue) ,XIO(SIC002.RunCommand) ONS(SIC002.StopOns) OTU(DigitalPoint[Address].CurrentValue) ];
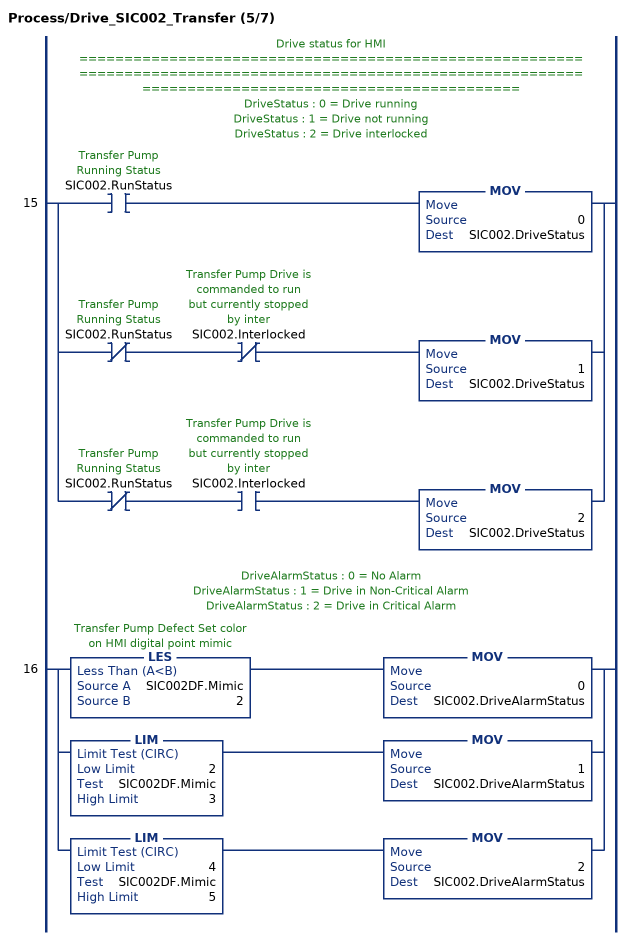
   // Drive status for HMI
   // ==========================================================================================================================================================
   //  DriveStatus : 0 = Drive running
   //  DriveStatus : 1 = Drive not running
   //  DriveStatus : 2 = Drive interlocked
   15: [XIC(SIC002.RunStatus) MOV(0,SIC002.DriveStatus) ,XIO(SIC002.RunStatus) XIO(SIC002.Interlocked) MOV(1,SIC002.DriveStatus) ,XIO(SIC002.RunStatus) XIC(SIC002.Interlocked) MOV(2,SIC002.DriveStatus) ];
   // DriveAlarmStatus : 0 = No Alarm
   //  DriveAlarmStatus : 1 = Drive in Non-Critical Alarm
   //  DriveAlarmStatus : 2 = Drive in Critical Alarm
   16: [LES(SIC002DF.Mimic,2) MOV(0,SIC002.DriveAlarmStatus) ,LIM(2,SIC002DF.Mimic,3) MOV(1,SIC002.DriveAlarmStatus) ,LIM(4,SIC002DF.Mimic,5) MOV(2,SIC002.DriveAlarmStatus) ];
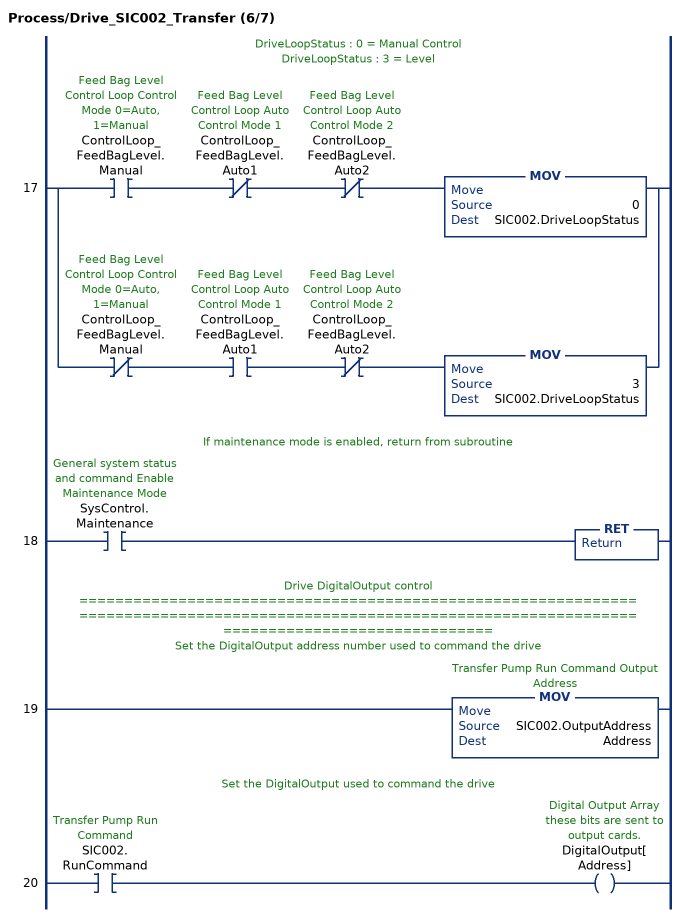
   // DriveLoopStatus : 0 = Manual Control
   //  DriveLoopStatus : 3 = Level
   17: [XIC(ControlLoop_FeedBagLevel.Manual) XIO(ControlLoop_FeedBagLevel.Auto1) XIO(ControlLoop_FeedBagLevel.Auto2) MOV(0,SIC002.DriveLoopStatus) ,XIO(ControlLoop_FeedBagLevel.Manual) XIC(ControlLoop_FeedBagLevel.Auto1) XIO(ControlLoop_FeedBagLevel.Auto2) MOV(3,SIC002.DriveLoopStatus) ];
   // If maintenance mode is enabled, return from subroutine
   18: XIC(SysControl.Maintenance)RET();
   // Drive DigitalOutput control
   // ==========================================================================================================================================================
   // Set the DigitalOutput address number used to command the drive
   19: MOV(SIC002.OutputAddress,Address);
   // Set the DigitalOutput used to command the drive
   20: XIC(SIC002.RunCommand)OTE(DigitalOutput[Address]);
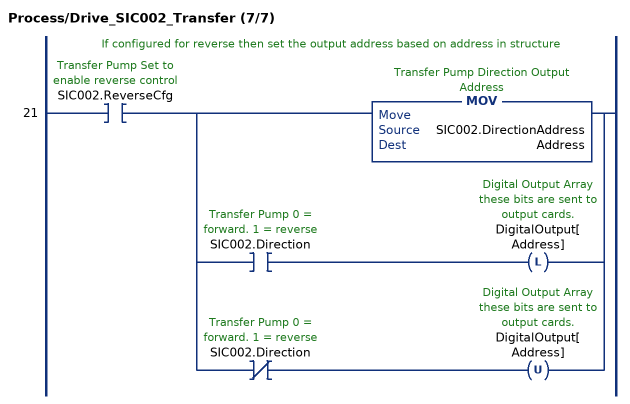
   // If configured for reverse then set the output address based on address in structure
   21: XIC(SIC002.ReverseCfg)[MOV(SIC002.DirectionAddress,Address) ,XIC(SIC002.Direction) OTL(DigitalOutput[Address]) ,XIO(SIC002.Direction) OTU(DigitalOutput[Address]) ];
END_ROUTINE
